TYPE ST_Actuator_HMI_Interface :
STRUCT
	HMIbaseDevice		: ST_Device_HMI_Interface; 
	stsActuated			: BOOL;
	ocmdActuate			: BOOL;
	ocmdReset			: BOOL;
	setActuate			: BOOL;
END_STRUCT
END_TYPE

(* stored: Version 1.1.0.1
   DUT ST_Actuator_HMI_Interface: Id {c487ca2e-f909-46b4-90db-25707195071a} *)
